(* PLC project g_ctd_load, Anonymous Benchmark Suite 1.0 *)
(* stored: creationDateTime 2026-08-26T00:00:00 *)

PROGRAM g_ctd_load
  VAR_INPUT
    Pulse : BOOL;
    Load : BOOL;
  END_VAR
  VAR_OUTPUT
    Empty : BOOL;
  END_VAR
  VAR
    CTD0 : CTD;
  END_VAR

(* LD diagram, written out as Structured Text *)
CTD0(CD := Pulse, PV := 2, LD := Load);
Empty := CTD0.Q;
END_PROGRAM

CONFIGURATION Config0
  RESOURCE Res0 ON PLC
    TASK tcyclic(INTERVAL := T#10ms, PRIORITY := 0);
    PROGRAM inst0 WITH tcyclic : g_ctd_load;
  END_RESOURCE
END_CONFIGURATION
